Fanuc KAREL source: KT00470.KL

PROGRAM KT00470
%NOLOCKGROUP
VAR
  P1: JOINTPOS
  P2: JOINTPOS
  OUT: BOOLEAN
BEGIN
  OUT = P1 >= P2
END KT00470
